(* IEC 61131-3 sources: llm-plc-st-eval/data/calibracion/qwen2.5-coder_14b/B1/zero_shot, 3 files *)

(* ---- ejec_1.st ---- *)
```pascal
FUNCTION_BLOCK FB_Motor
VAR_INPUT
    btnMarcha : BOOL;  // Botón de marcha
    btnParo : BOOL;    // Botón de paro
    btnEmerg : BOOL;   // Botón de paro de emergencia
END_VAR

VAR_OUTPUT
    motorOn : BOOL;    // Estado del motor (encendido/apagado)
END_VAR

VAR
    emergenciaActiva : BOOL := FALSE;  // Bandera para indicar si hay una parada de emergencia
END_VAR

// Programa principal
IF btnEmerg THEN
    // Si se activa el botón de emergencia, detener el motor y activar la bandera de emergencia
    motorOn := FALSE;
    emergenciaActiva := TRUE;
ELSIF emergenciaActiva THEN
    // Si hay una parada de emergencia activa, mantener el motor apagado
    motorOn := FALSE;
ELSIF btnParo THEN
    // Si se presiona el botón de paro, detener el motor
    motorOn := FALSE;
ELSIF btnMarcha THEN
    // Si se presiona el botón de marcha, encender el motor
    motorOn := TRUE;
END_IF;
```

(* ---- ejec_2.st ---- *)
```pascal
FUNCTION_BLOCK FB_Motor
VAR_INPUT
    btnMarcha : BOOL; // Botón de marcha
    btnParo : BOOL; // Botón de paro
    btnEmerg : BOOL; // Botón de emergencia
END_VAR

VAR_OUTPUT
    motorOn : BOOL; // Estado del motor
END_VAR

VAR
    estadoEmergencia : BOOL := FALSE; // Bandera de emergencia
END_VAR

// Programa principal
IF btnEmerg THEN
    // Si se presiona el botón de emergencia
    estadoEmergencia := TRUE;
    motorOn := FALSE; // Apaga el motor
ELSIF estadoEmergencia THEN
    // Si hay una emergencia activa, no se permite el arranque
    motorOn := FALSE;
ELSIF btnParo THEN
    // Si se presiona el botón de paro
    motorOn := FALSE; // Apaga el motor
ELSIF btnMarcha THEN
    // Si se presiona el botón de marcha
    motorOn := TRUE; // Enciende el motor
END_IF;
```

Este código implementa un control de arranque y paro de un motor trifásico siguiendo las especificaciones proporcionadas. El motor se encenderá cuando se presione el botón de marcha y permanecerá encendido incluso al soltar el botón. El motor se apagará cuando se presione el botón de paro o el botón de emergencia. Después de un paro de emergencia, el motor no se podrá arrancar aunque el botón de marcha esté pulsado.

(* ---- ejec_3.st ---- *)
```pascal
FUNCTION_BLOCK FB_Motor
VAR_INPUT
    btnMarcha : BOOL; // Botón de marcha
    btnParo : BOOL; // Botón de paro
    btnEmerg : BOOL; // Botón de emergencia
END_VAR

VAR_OUTPUT
    motorOn : BOOL; // Estado del motor (encendido/apagado)
END_VAR

VAR
    emergenciaActiva : BOOL := FALSE; // Estado de emergencia activa
END_VAR

// Programa principal
IF btnEmerg THEN
    emergenciaActiva := TRUE; // Activar estado de emergencia
    motorOn := FALSE; // Apagar motor en caso de emergencia
ELSIF emergenciaActiva THEN
    motorOn := FALSE; // Mantener motor apagado si hay emergencia activa
ELSE
    IF btnParo THEN
        motorOn := FALSE; // Apagar motor si se presiona el botón de paro
    ELSE
        motorOn := btnMarcha; // Mantener motor encendido si se mantiene presionado el botón de marcha
    END_IF
END_IF;
```

Este código implementa un control de arranque y paro de un motor trifásico siguiendo las especificaciones proporcionadas. El motor se encenderá cuando se presione el botón de marcha y se mantendrá encendido mientras se mantenga presionado. El motor se apagará cuando se presione el botón de paro o el botón de emergencia. Después de un paro de emergencia, el motor no se podrá volver a encender aunque se mantenga presionado el botón de marcha.
